Fanuc KAREL source: kt00493.KL

-- PROVISIONAL review KL for V1013-1; original PC SHA256 1a2c18b978e91ae4f8c5737863204241e86155860bd9376f604521f73ae2bddc
-- Incomplete behavior may be omitted. Consult companion uncertainty JSON. Do not deploy.
PROGRAM KT00493
%NOLOCKGROUP
VAR
  OUT : BOOLEAN
-- UNRESOLVED_DECL P1 type=000102
-- UNRESOLVED_DECL P2 type=000101
BEGIN
  -- UNRESOLVED_PC offsets 5-20; opcodes 2E,22,32,35
  -- UNRESOLVED_PC offsets 25-53; opcodes 49,7E,49,AC,23
  -- UNRESOLVED_PC offsets 58-62; opcodes 7F
END KT00493
